FUNCTION_BLOCK PUMP_STATION_SUPERVISOR (* Migrated from IEC 61131-3 ST *)
  (* Standard: 61499-2 *)
  (* Version 1.0, 2026-11-06, st2fb *)
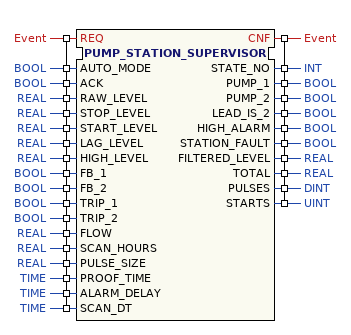
  EVENT_INPUT
    REQ WITH AUTO_MODE, ACK, RAW_LEVEL, STOP_LEVEL, START_LEVEL, LAG_LEVEL, HIGH_LEVEL, FB_1, FB_2, TRIP_1, TRIP_2, FLOW, SCAN_HOURS, PULSE_SIZE, PROOF_TIME, ALARM_DELAY, SCAN_DT;
  END_EVENT
  EVENT_OUTPUT
    CNF WITH STATE_NO, PUMP_1, PUMP_2, LEAD_IS_2, HIGH_ALARM, STATION_FAULT, FILTERED_LEVEL, TOTAL, PULSES, STARTS;
  END_EVENT
  VAR_INPUT
    AUTO_MODE : BOOL;
    ACK : BOOL;
    RAW_LEVEL : REAL;
    STOP_LEVEL : REAL;
    START_LEVEL : REAL;
    LAG_LEVEL : REAL;
    HIGH_LEVEL : REAL;
    FB_1 : BOOL;
    FB_2 : BOOL;
    TRIP_1 : BOOL;
    TRIP_2 : BOOL;
    FLOW : REAL;
    SCAN_HOURS : REAL;
    PULSE_SIZE : REAL;
    PROOF_TIME : TIME;
    ALARM_DELAY : TIME;
    SCAN_DT : TIME;
  END_VAR
  VAR_OUTPUT
    STATE_NO : INT;
    PUMP_1 : BOOL;
    PUMP_2 : BOOL;
    LEAD_IS_2 : BOOL;
    HIGH_ALARM : BOOL;
    STATION_FAULT : BOOL;
    FILTERED_LEVEL : REAL;
    TOTAL : REAL;
    PULSES : DINT;
    STARTS : UINT;
  END_VAR
  VAR
    FAILED_1_Q1 : BOOL := FALSE;
    FAILED_2_Q1 : BOOL := FALSE;
    PROOF_TIMER_IN : BOOL := FALSE;
    PROOF_TIMER_PT : TIME := T#0s;
    PROOF_TIMER_Q : BOOL := FALSE;
    PROOF_TIMER_ET : TIME := T#0s;
    PROOF_TIMER_STATE : INT := 0;
    PROOF_TIMER_PREV_IN : BOOL := FALSE;
    PROOF_TIMER_START_TIME : TIME := T#0s;
    ALARM_TIMER_IN : BOOL := FALSE;
    ALARM_TIMER_PT : TIME := T#0s;
    ALARM_TIMER_Q : BOOL := FALSE;
    ALARM_TIMER_ET : TIME := T#0s;
    ALARM_TIMER_STATE : INT := 0;
    ALARM_TIMER_PREV_IN : BOOL := FALSE;
    ALARM_TIMER_START_TIME : TIME := T#0s;
    ACK_EDGE_CLK : BOOL := FALSE;
    ACK_EDGE_Q : BOOL := FALSE;
    ACK_EDGE_M : BOOL := FALSE;
    PASSES : INT := 0;
    I : INT := 0;
    STEP_SIZE : REAL := 0.0;
    PENDING : REAL := 0.0;
    LEAD_RUNNING_FB : BOOL := FALSE;
    LEAD_FAILED : BOOL := FALSE;
    LAG_FAILED : BOOL := FALSE;
    ST2FB_NOW : TIME := T#0s;
  END_VAR
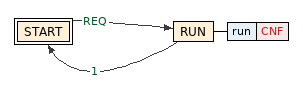
  EC_STATES
    START;
    RUN : run -> CNF;
  END_STATES
  EC_TRANSITIONS
    START TO RUN := REQ;
    RUN TO START := 1;
  END_TRANSITIONS
  ALGORITHM run IN ST:
ST2FB_NOW := ST2FB_NOW + SCAN_DT;
STEP_SIZE := RAW_LEVEL - FILTERED_LEVEL;
IF (STEP_SIZE > 1.0) OR (STEP_SIZE < -1.0) THEN
  PASSES := 4;
ELSE
  PASSES := 1;
END_IF;
FOR I := 1 TO PASSES DO
  FILTERED_LEVEL := FILTERED_LEVEL + 0.25 * (RAW_LEVEL - FILTERED_LEVEL);
END_FOR;

ACK_EDGE_CLK := ACK;
ACK_EDGE_Q := ACK_EDGE_CLK AND NOT ACK_EDGE_M;
ACK_EDGE_M := ACK_EDGE_CLK;

FAILED_1_Q1 := (TRIP_1 OR (PROOF_TIMER_Q AND NOT LEAD_IS_2)) OR (NOT ACK_EDGE_Q AND FAILED_1_Q1);
FAILED_2_Q1 := (TRIP_2 OR (PROOF_TIMER_Q AND LEAD_IS_2)) OR (NOT ACK_EDGE_Q AND FAILED_2_Q1);
IF LEAD_IS_2 THEN
  LEAD_FAILED := FAILED_2_Q1;
  LAG_FAILED := FAILED_1_Q1;
  LEAD_RUNNING_FB := FB_2;
ELSE
  LEAD_FAILED := FAILED_1_Q1;
  LAG_FAILED := FAILED_2_Q1;
  LEAD_RUNNING_FB := FB_1;
END_IF;

IF NOT AUTO_MODE AND STATE_NO <> 5 THEN
  STATE_NO := 0;
END_IF;
CASE STATE_NO OF
  0:
    IF AUTO_MODE THEN
      STATE_NO := 1;
    END_IF;
  1:
    IF LEAD_FAILED AND LAG_FAILED THEN
      STATE_NO := 5;
    ELSIF LEAD_FAILED THEN
      LEAD_IS_2 := NOT LEAD_IS_2;
    ELSIF FILTERED_LEVEL >= START_LEVEL THEN
      STARTS := STARTS + 1;
      STATE_NO := 2;
    END_IF;
  2:
    IF LEAD_FAILED THEN
      STATE_NO := 1;
    ELSIF LEAD_RUNNING_FB THEN
      STATE_NO := 3;
    END_IF;
  3:
    IF LEAD_FAILED THEN
      STATE_NO := 1;
    ELSIF FILTERED_LEVEL <= STOP_LEVEL THEN
      LEAD_IS_2 := NOT LEAD_IS_2;
      STATE_NO := 1;
    ELSIF (FILTERED_LEVEL >= LAG_LEVEL) AND NOT LAG_FAILED THEN
      STATE_NO := 4;
    END_IF;
  4:
    IF LEAD_FAILED THEN
      STATE_NO := 1;
    ELSIF LAG_FAILED OR (FILTERED_LEVEL < LAG_LEVEL) THEN
      STATE_NO := 3;
    END_IF;
  5:
    IF NOT (LEAD_FAILED OR LAG_FAILED) THEN
      STATE_NO := 0;
    END_IF;
ELSE
  STATE_NO := 0;
END_CASE;

PROOF_TIMER_IN := (STATE_NO = 2) AND NOT LEAD_RUNNING_FB;
PROOF_TIMER_PT := PROOF_TIME;
IF (PROOF_TIMER_STATE = 0) AND NOT PROOF_TIMER_PREV_IN AND PROOF_TIMER_IN THEN
  PROOF_TIMER_STATE := 1;
  PROOF_TIMER_Q := FALSE;
  PROOF_TIMER_START_TIME := ST2FB_NOW;
ELSE
  IF NOT PROOF_TIMER_IN THEN
    PROOF_TIMER_ET := T#0s;
    PROOF_TIMER_Q := FALSE;
    PROOF_TIMER_STATE := 0;
  ELSIF PROOF_TIMER_STATE = 1 THEN
    IF PROOF_TIMER_START_TIME + PROOF_TIMER_PT <= ST2FB_NOW THEN
      PROOF_TIMER_STATE := 2;
      PROOF_TIMER_Q := TRUE;
      PROOF_TIMER_ET := PROOF_TIMER_PT;
    ELSE
      PROOF_TIMER_ET := ST2FB_NOW - PROOF_TIMER_START_TIME;
    END_IF;
  END_IF;
END_IF;
PROOF_TIMER_PREV_IN := PROOF_TIMER_IN;

STATION_FAULT := STATE_NO = 5;

IF (STATE_NO >= 2) AND (STATE_NO <= 4) THEN
  PUMP_1 := NOT LEAD_IS_2 OR (STATE_NO = 4);
  PUMP_2 := LEAD_IS_2 OR (STATE_NO = 4);
ELSE
  PUMP_1 := FALSE;
  PUMP_2 := FALSE;
END_IF;

ALARM_TIMER_IN := FILTERED_LEVEL >= HIGH_LEVEL;
ALARM_TIMER_PT := ALARM_DELAY;
IF (ALARM_TIMER_STATE = 0) AND NOT ALARM_TIMER_PREV_IN AND ALARM_TIMER_IN THEN
  ALARM_TIMER_STATE := 1;
  ALARM_TIMER_Q := FALSE;
  ALARM_TIMER_START_TIME := ST2FB_NOW;
ELSE
  IF NOT ALARM_TIMER_IN THEN
    ALARM_TIMER_ET := T#0s;
    ALARM_TIMER_Q := FALSE;
    ALARM_TIMER_STATE := 0;
  ELSIF ALARM_TIMER_STATE = 1 THEN
    IF ALARM_TIMER_START_TIME + ALARM_TIMER_PT <= ST2FB_NOW THEN
      ALARM_TIMER_STATE := 2;
      ALARM_TIMER_Q := TRUE;
      ALARM_TIMER_ET := ALARM_TIMER_PT;
    ELSE
      ALARM_TIMER_ET := ST2FB_NOW - ALARM_TIMER_START_TIME;
    END_IF;
  END_IF;
END_IF;
ALARM_TIMER_PREV_IN := ALARM_TIMER_IN;
HIGH_ALARM := ALARM_TIMER_Q;

IF PUMP_1 OR PUMP_2 THEN
  TOTAL := TOTAL + FLOW * SCAN_HOURS;
  PENDING := PENDING + FLOW * SCAN_HOURS;
  WHILE PENDING >= PULSE_SIZE DO
    PENDING := PENDING - PULSE_SIZE;
    PULSES := PULSES + 1;
  END_WHILE;
END_IF;
  END_ALGORITHM
END_FUNCTION_BLOCK
